(* IEC 61131-3 sources: tsplc/packages/vscode-extension/tests/fixtures/conveyor, 1 file *)

(* ---- Main.st ---- *)
PROGRAM Main
VAR
	Inbound : FB_Conveyor;
END_VAR

Inbound(Conveyor := PlantIO.Inbound);
Inbound.SetMotionSignal(Asserted := TRUE);
END_PROGRAM
